// TIA Portal V20 export
Screen "15_SubMenus_ProductionData"  100x768
  ScreenItem "txtOverview_15" at -1,713 size 100x53  Type=HmiTextBox
  ScreenItem "txtOverview_1" at -1,653 size 100x52  Type=HmiTextBox
  ScreenItem "txtOverview_2" at -1,593 size 100x52  Type=HmiTextBox
  ScreenItem "txtOverview_3" at -1,533 size 100x52  Type=HmiTextBox
  ScreenItem "txtOverview_4" at -1,473 size 100x52  Type=HmiTextBox
  ScreenItem "txtOverview_5" at -1,413 size 100x52  Type=HmiTextBox
  ScreenItem "txtOverview_6" at -1,353 size 100x52  Type=HmiTextBox
  ScreenItem "txtOverview_7" at -1,293 size 100x52  Type=HmiTextBox
  ScreenItem "txtOverview_8" at -1,233 size 100x52  Type=HmiTextBox
  ScreenItem "txtOverview_9" at -1,173 size 100x52  Type=HmiTextBox
  ScreenItem "txtOverview_10" at -1,113 size 100x52  Type=HmiTextBox
  ScreenItem "txtOverview_11" at -1,53 size 100x52  Type=HmiTextBox
  ScreenItem "txtOverview_12" at -1,-7 size 100x52  Type=HmiTextBox
  ScreenItem "线_1" at 1,409 size 97x0  Type=HmiLine
